(* IEC 61131-3 sources: codesys-framework/txt/application/ToDo/Hardware/IO/Camera/FB_Camera/Public, 8 files *)

(* ---- Connect.method.st ---- *)
METHOD Connect : BOOL
VAR_INPUT
END_VAR

// --- BEGIN IMPLEMENTATION ---

IF _xDone  THEN
	Connect := TRUE;
	RETURN;
END_IF

IF _eState = E_CameraStates.Standby THEN
	_eState := E_CameraStates.Connect;
END_IF

(* ---- Disconnect.method.st ---- *)
METHOD Disconnect : BOOL
VAR_INPUT
END_VAR

// --- BEGIN IMPLEMENTATION ---

IF _xDone  THEN
	Disconnect := TRUE;
	RETURN;
END_IF

IF _eState = E_CameraStates.Standby THEN
	_eState := E_CameraStates.Disconnect;
END_IF

(* ---- GetResult.method.st ---- *)
METHOD GetResult : STRING(255)
VAR_INPUT
END_VAR

// --- BEGIN IMPLEMENTATION ---

GetResult := _sResult;

(* ---- Initialize.method.st ---- *)
METHOD Initialize
VAR_INPUT
END_VAR

// --- BEGIN IMPLEMENTATION ---

_xBusy := FALSE;
_xDone := FALSE;
_xError := FALSE;
_iErrorId := 0;
_sError := '';
_xConnected := FALSE;
_iStateMonitor := 0;
_iStateConnect := 0;
_iStateSetJob := 0;
_iStateTakePicture := 0;
_iStateConnectMethod := 0;
_iStateDisconnect := 0;

_sFeedBack := '';
_sJob := '';
_sPicture := '';
_id := 0;

_tonPicture.IN := FALSE;
_write.xExecute := FALSE;
_tonSelectJob.IN := FALSE;

_eState := E_CameraStates.Connect;

(* ---- Reset.method.st ---- *)
METHOD Reset
VAR_INPUT
END_VAR

// --- BEGIN IMPLEMENTATION ---

_xBusy := FALSE;
_xDone := FALSE;
_xError := FALSE;
_iErrorId := 0;
_sError := '';
_xConnected := FALSE;
_iStateMonitor := 0;
_iStateConnect := 0;
_iStateConnectMethod := 0;
_iStateSetJob := 0;
_iStateTakePicture := 0;

_sFeedBack := '';
_sJob := '';
_sPicture := '';
_id := 0;

_write.xExecute := FALSE;

_clientRead.xEnable := FALSE;
_clientWrite.xEnable := FALSE;

(* ---- ResetResult.method.st ---- *)
METHOD ResetResult
VAR_INPUT
END_VAR

// --- BEGIN IMPLEMENTATION ---

_sResultPrev := _sResult;
_sResult := '';

(* ---- SetJob.method.st ---- *)
METHOD SetJob : BOOL
VAR_INPUT
	id 		: UINT;
END_VAR

// --- BEGIN IMPLEMENTATION ---

IF _xDone  THEN
	SetJob := TRUE;
	RETURN;
END_IF

IF _eState = E_CameraStates.Standby THEN
	_id := id;
	_eState := E_CameraStates.SelectJob;
END_IF

(* ---- TakePicture.method.st ---- *)
METHOD TakePicture : BOOL
VAR_INPUT
	pictureId		: STRING;
END_VAR
VAR
	dataLength		: INT := 0;
	sDataLength		: STRING;
	operationInst	: STRING := 'TRX';
END_VAR

// --- BEGIN IMPLEMENTATION ---

dataLength := LEN(pictureId);
sDataLength := INT_TO_STRING(dataLength);

WHILE LEN(sDataLength) < 2 DO
	sDataLength := CONCAT('0', INT_TO_STRING(dataLength));
END_WHILE

_sPictureId := 	CONCAT(operationInst,
					CONCAT(sDataLength, pictureId)
				);

IF _xDone  THEN
	TakePicture := TRUE;
	RETURN;
END_IF

IF _eState = E_CameraStates.Standby THEN
	_eState := E_CameraStates.TakePicture;
END_IF
